PROGRAM main
  VAR
    Fill_Btn AT %IX0.0 : BOOL;
    Disch_Btn AT %IX0.1 : BOOL;
    Fill_Valve AT %QX0.0 : BOOL;
    Disch_Valve AT %QX0.1 : BOOL;
    T_Fill : TON;
    T_Disch : TON;
    Fill_Seq : BOOL;
    Disch_Seq : BOOL;
    Fill_Light AT %QX0.2 : BOOL;
    Timer_Disp AT %QW0 : INT;
    Disch_Light AT %QX0.3 : BOOL;
    Fill_sec : LREAL;
    Left_Calc : LREAL;
    Disch_sec : LREAL;
  END_VAR
  VAR_EXTERNAL
  END_VAR
  VAR_INPUT
  END_VAR

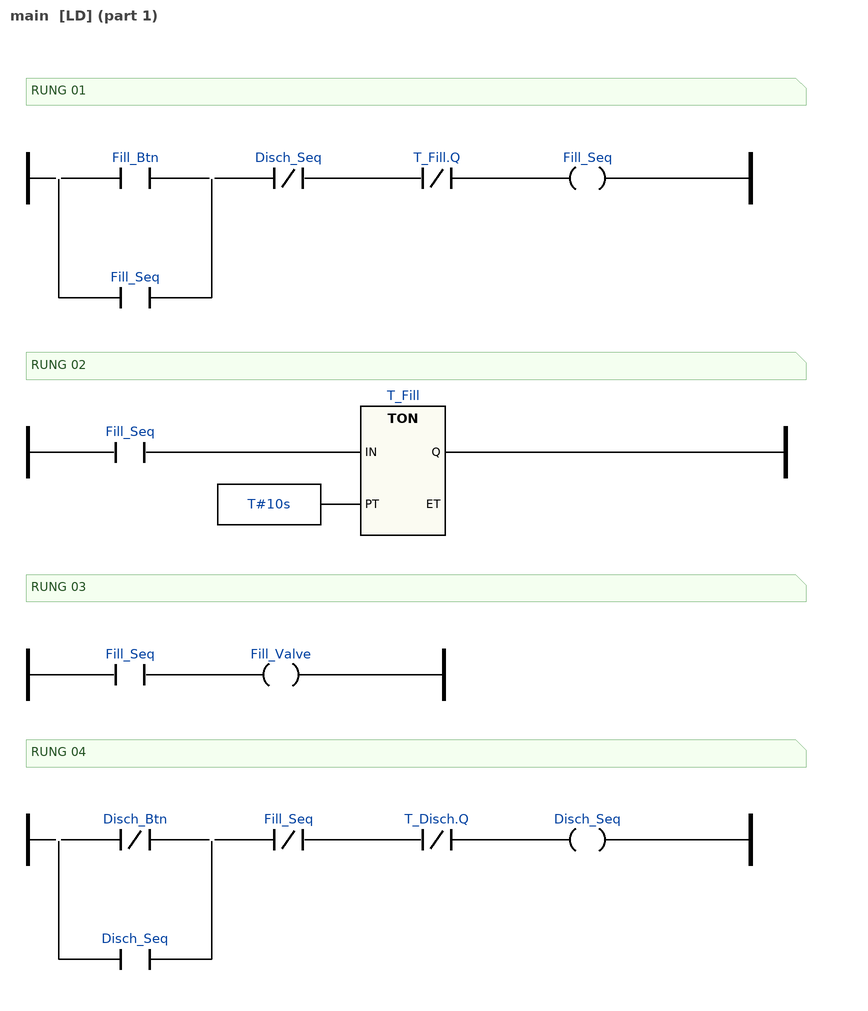
(* LD diagram, written out as Structured Text *)
(* RUNG 01 *)
Fill_Seq := (Fill_Btn OR Fill_Seq) AND NOT Disch_Seq AND NOT T_Fill.Q;
(* RUNG 02 *)
(* RUNG 03 *)
Fill_Valve := Fill_Seq;
(* RUNG 04 *)
Disch_Seq := (Disch_Seq OR NOT Disch_Btn) AND NOT Fill_Seq AND NOT T_Disch.Q;
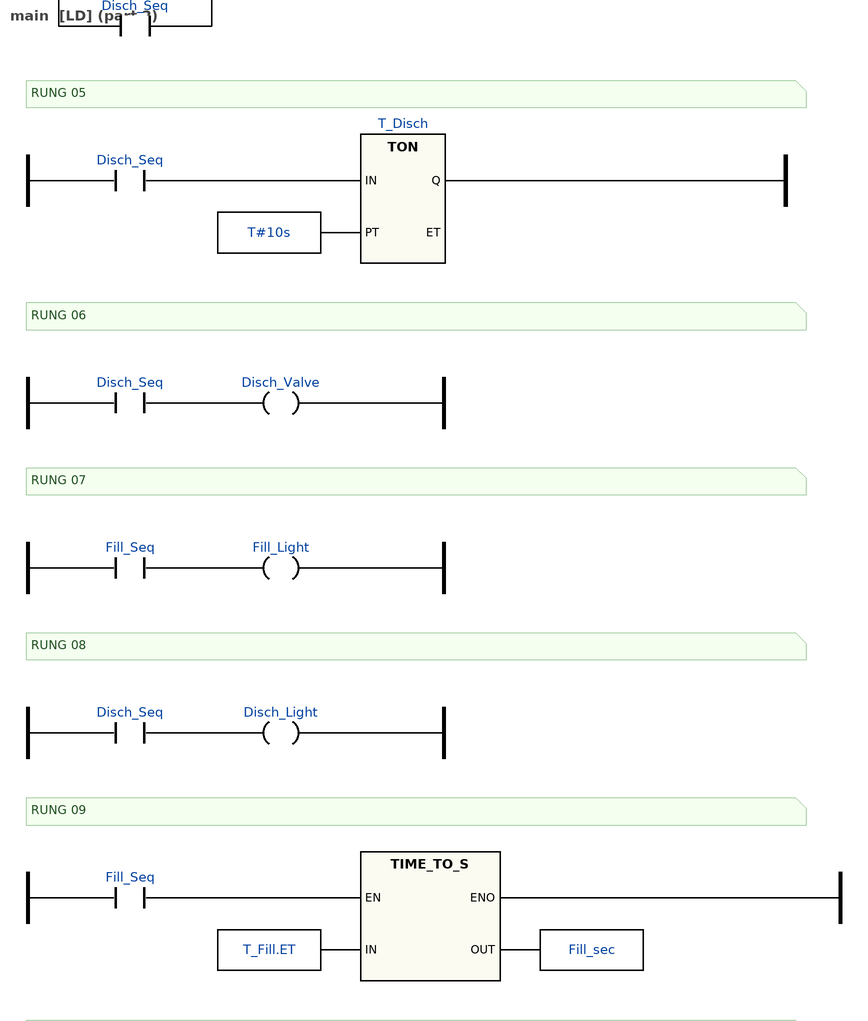
(* RUNG 05 *)
(* RUNG 06 *)
Disch_Valve := Disch_Seq;
(* RUNG 07 *)
Fill_Light := Fill_Seq;
(* RUNG 08 *)
Disch_Light := Disch_Seq;
(* RUNG 09 *)
IF Fill_Seq THEN Fill_sec := TIME_TO_S(T_Fill.ET); END_IF;
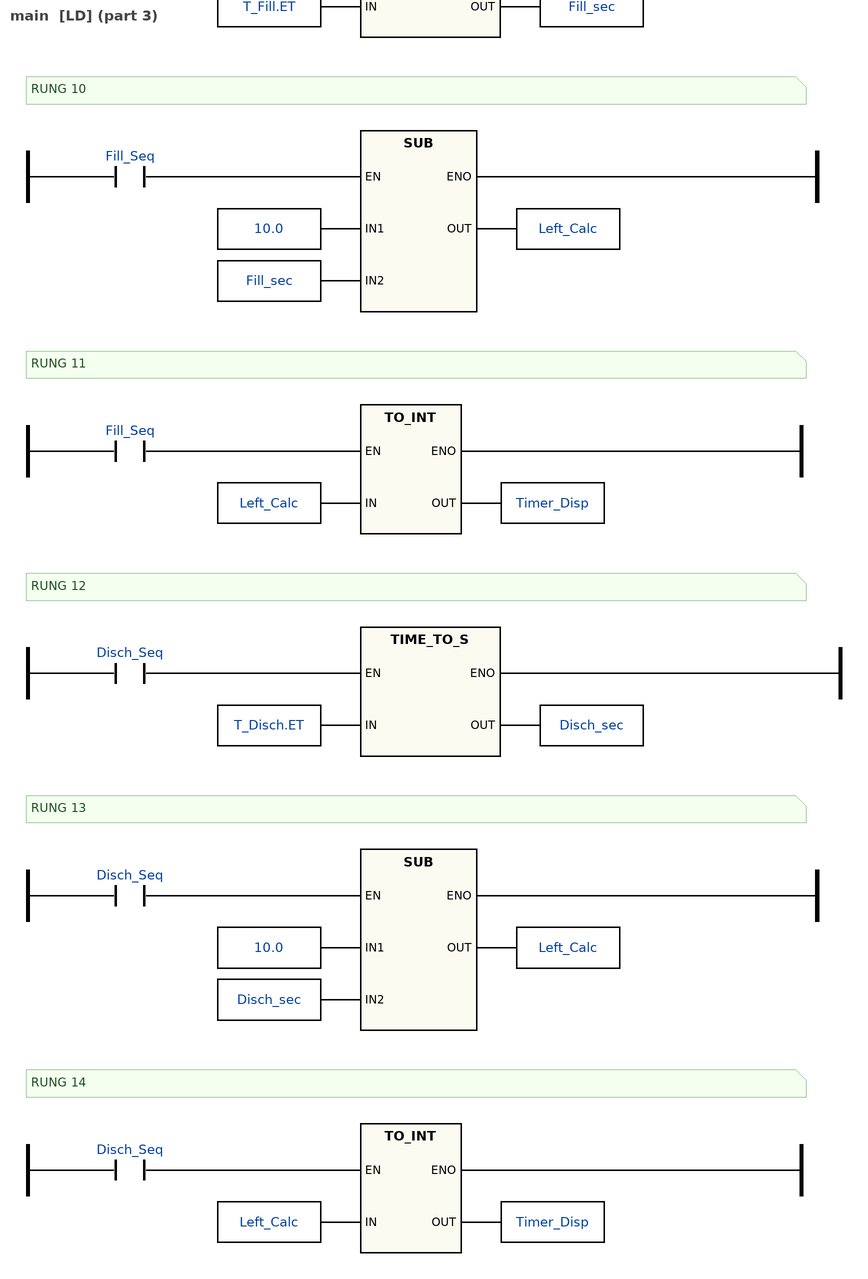
(* RUNG 10 *)
IF Fill_Seq THEN Left_Calc := 10.0 - Fill_sec; END_IF;
(* RUNG 11 *)
IF Fill_Seq THEN Timer_Disp := TO_INT(Left_Calc); END_IF;
(* RUNG 12 *)
IF Disch_Seq THEN Disch_sec := TIME_TO_S(T_Disch.ET); END_IF;
(* RUNG 13 *)
IF Disch_Seq THEN Left_Calc := 10.0 - Disch_sec; END_IF;
(* RUNG 14 *)
IF Disch_Seq THEN Timer_Disp := TO_INT(Left_Calc); END_IF;
T_Fill(IN := Fill_Seq, PT := T#10s);
T_Disch(IN := Disch_Seq, PT := T#10s);
END_PROGRAM
